(* IEC 61131-3 sources: ayran-mini-fabrika/plc/build (part 7) *)

  CASE STP OF
    0:  (* idle *)
      WANT := WORD#0;
      PUMP_REQ := FALSE;
      IF NOT WAIT_START AND (ALARMS AND ALARM_MASK) = WORD#0 THEN
        IF CIP_REQ THEN
          CIP_REQ := FALSE;
          STP := 40;
        ELSIF REQ AND NOT CIP_DUE AND NOT DI_T1_LOW THEN
          BATCH := 0;
          IF LINE_PRODUCT THEN STP := 10; ELSE STP := 20; END_IF;
        END_IF;
      END_IF;

    20: (* fill the line with product: first liquid to the drain *)
      WANT := WORD#16#0022;            (* V_PROD + V_DRAIN *)
      PUMP_REQ := TRUE;
      IF T_INWIN.Q THEN
        LINE_PRODUCT := TRUE;
        STP := 10;                     (* the route manager stops the pump and changes the route *)
      ELSIF STEP_SCANS > 2250 THEN
        ALARMS := ALARMS OR WORD#16#0200;   (* product conductivity not detected within 45 s *)
      END_IF;

    10: (* transfer to the filling tank *)
      WANT := WORD#16#0012;            (* V_PROD + V_FILL *)
      PUMP_REQ := TRUE;
      IF T_FOREIGN.Q THEN
        LINE_PRODUCT := FALSE;
        ALARMS := ALARMS OR WORD#16#0004;
      ELSIF NOT REQ OR DI_T1_LOW OR SINCE >= CIP_LIMIT OR CIP_REQ THEN
        STP := 0;
      END_IF;

    40: (* CIP preparation: empty route for the line, prove all valves closed *)
      WANT := WORD#0;
      PUMP_REQ := FALSE;
      LINE_PRODUCT := FALSE;
      CAUSTIC_IN := FALSE;
      CIP_SCANS := 0;
      MIN_T := 32000;
      MIN_F := 32000;
      FINAL_COND := 0;
      IF IW_CIP_LVL < CIP_LVL_MIN THEN
        ALARMS := ALARMS OR WORD#16#0100;
      ELSIF RSTATE = 0 AND ROUTE_OK THEN
        STP := 41;
      END_IF;

    41: (* wait for the caustic temperature *)
      WANT := WORD#0;
      PUMP_REQ := FALSE;
      IF IW_CIP_T >= CAUSTIC_SP - 50 THEN
        STP := 42;
      ELSIF STEP_TO THEN
        ALARMS := ALARMS OR WORD#16#0080;
      END_IF;

    42: (* pre-rinse: water to the drain *)
      WANT := WORD#16#0024;            (* V_WATER + V_DRAIN *)
      PUMP_REQ := TRUE;
      IF VOL >= RINSE_KG THEN
        WATER_REF := IW_COND;           (* conductivity of the inlet water: the criterion for the final rinse *)
        STP := 43;
      ELSIF STEP_TO THEN
        ALARMS := ALARMS OR WORD#16#0080;
      END_IF;

    43: (* caustic: first to the drain, to the caustic tank once caustic arrives (phase separation) *)
      PUMP_REQ := TRUE;
      IF NOT CAUSTIC_IN AND RSTATE = 0 AND IW_COND >= COND_CAUSTIC THEN CAUSTIC_IN := TRUE; END_IF;
      IF CAUSTIC_IN THEN
        WANT := WORD#16#0048;          (* V_CAUSTIC + V_CIPRET *)
      ELSE
        WANT := WORD#16#0028;          (* V_CAUSTIC + V_DRAIN *)
      END_IF;
      (* CIP record: the lowest values in the counted hold window *)
      IF HOLD_OK THEN
        IF IW_RET_T < MIN_T THEN MIN_T := IW_RET_T; END_IF;
        IF IW_FLOW < MIN_F THEN MIN_F := IW_FLOW; END_IF;
      ELSE
        MIN_T := 32000;
        MIN_F := 32000;
      END_IF;
      IF T_HOLD.Q THEN
        STP := 44;
      ELSIF STEP_TO THEN
        ALARMS := ALARMS OR WORD#16#0080;
      END_IF;

    44: (* final rinse: until no caustic is left *)
      WANT := WORD#16#0024;
      PUMP_REQ := TRUE;
      IF VOL >= RINSE_KG AND IW_COND <= WATER_REF + RINSE_MARGIN THEN
        FINAL_COND := IW_COND;
        STP := 45;
      ELSIF STEP_TO THEN
        ALARMS := ALARMS OR WORD#16#0080;
      END_IF;

    45: (* completed *)
      WANT := WORD#0;
      PUMP_REQ := FALSE;
      SINCE := 0;
      CIP_DUE := FALSE;
      ABORT_WARN := FALSE;
      CIP_RES := 1;
      CIP_DUR := CIP_SCANS / 50;
      STP := 0;
  END_CASE;
  IF STP >= 40 AND STP <= 44 AND CIP_SCANS < 30000 THEN CIP_SCANS := CIP_SCANS + 1; END_IF;
  IF CIP_RES = 2 OR CIP_RES = 3 THEN CIP_DUR := CIP_SCANS / 50; END_IF;

  (* =================== 4. Route manager =================== *)
  IF (ALARMS AND ALARM_MASK) <> WORD#0 THEN WANT := WORD#0; END_IF;
  IF WANT <> CUR AND RSTATE = 0 THEN RSTATE := 1; END_IF;
  T_ROUTE(IN := RSTATE = 1, PT := T#3s);
  T_STROKE(IN := RSTATE = 2, PT := T#1s);
  IF RSTATE = 1 THEN
    VALVES := CUR AND WANT;            (* close the ones not in the new route *)
    IF ((NOT WANT) AND WORD#16#007E AND (NOT CLOSED)) = WORD#0 THEN
      RSTATE := 2;
    ELSIF T_ROUTE.Q THEN
      ALARMS := ALARMS OR WORD#16#0008;
      RSTATE := 0;
      CUR := CUR AND WANT;
    END_IF;
  ELSIF RSTATE = 2 THEN
    VALVES := WANT;
    IF T_STROKE.Q THEN CUR := WANT; RSTATE := 0; END_IF;
  ELSE
    VALVES := CUR;
  END_IF;

  Q_P1 := PUMP_REQ AND RSTATE = 0 AND CUR = WANT AND CUR <> WORD#0 AND ROUTE_OK
          AND (ALARMS AND ALARM_MASK) = WORD#0;

  (* caustic tank thermostat (+/- 2 C), level and over-temperature interlock *)
  IF NOT ESTOP_OK OR IW_CIP_LVL < CIP_LVL_MIN OR IW_CIP_T > CAUSTIC_MAX THEN
    Q_HEAT := FALSE;
  ELSIF IW_CIP_T < CAUSTIC_SP - 20 THEN
    Q_HEAT := TRUE;
  ELSIF IW_CIP_T > CAUSTIC_SP + 20 THEN
    Q_HEAT := FALSE;
  END_IF;

  (* =================== 5. Outputs =================== *)
  WARNS := WORD#0;
  IF DI_T1_LOW THEN WARNS := WARNS OR WORD#16#0400; END_IF;
  IF CIP_DUE THEN WARNS := WARNS OR WORD#16#0800; END_IF;
  IF ABORT_WARN THEN WARNS := WARNS OR WORD#16#1000; END_IF;

  QW_DO := VALVES AND WORD#16#007E;
  IF Q_P1 THEN QW_DO := QW_DO OR WORD#16#0001; END_IF;
  IF Q_HEAT THEN QW_DO := QW_DO OR WORD#16#0080; END_IF;
  IF STP >= 40 THEN QW_DO := QW_DO OR WORD#16#0100; END_IF;

  IF (ALARMS AND WORD#16#0001) <> WORD#0 THEN
    QW_STATE := 11;
  ELSIF (ALARMS AND ALARM_MASK) <> WORD#0 THEN
    QW_STATE := 10;
  ELSIF STP = 0 AND CIP_DUE THEN
    QW_STATE := 9;
  ELSIF STP = 0 THEN
    QW_STATE := 0;
  ELSIF (STP = 10 OR STP = 20) AND RSTATE <> 0 THEN
    QW_STATE := 3;
  ELSIF STP = 10 THEN
    QW_STATE := 1;
  ELSIF STP = 20 THEN
    QW_STATE := 2;
  ELSE
    QW_STATE := STP - 36;             (* 40..44 -> 4..8 *)
  END_IF;

  QW_ALARM    := ALARMS OR WARNS;
  QW_STEP_T   := STEP_SCANS / 50;
  QW_SINCE    := SINCE;
  QW_BATCH    := BATCH;
  QW_CIP_RES  := CIP_RES;
  IF MIN_T = 32000 THEN QW_CIP_MINT := 0; ELSE QW_CIP_MINT := MIN_T; END_IF;
  IF MIN_F = 32000 THEN QW_CIP_MINF := 0; ELSE QW_CIP_MINF := MIN_F; END_IF;
  QW_CIP_COND := FINAL_COND;
  QW_CIP_DUR  := CIP_DUR;
  TRANSFERRING := STP = 10 AND Q_P1;
  QW_STATUS := WORD#0;
  IF WAIT_START THEN QW_STATUS := WORD#16#0080; END_IF;
  IF WAIT_START OR NOT IO_READY THEN
    QW_DO := WORD#0;
    Q_HEAT := FALSE; Q_P1 := FALSE;
  END_IF;
END_FUNCTION_BLOCK

PROGRAM Proses
  VAR
    (* --- blok 0: Fabrika --- *)
    FAB_IW_DI        AT %IW100 : WORD;  (* Fabrika paneli girisleri (bit paketli) *)
    FAB_IW_MAPVER    AT %IW101 : INT;  (* Sinyal haritasi surumu *)
    FAB_IW_SIM_HB    AT %IW102 : INT;  (* Simulator kalp atisi (100 ms) *)
    FAB_QW_DO        AT %QW100 : WORD;  (* Fabrika cikislari (bit paketli) *)
    FAB_QW_PLC_HB    AT %QW101 : INT;  (* Proses PLC (ya da tek PLC) kalp atisi (her tarama) *)
    FAB_QW_STATE     AT %QW102 : INT;  (* Fabrika durumu *)
    FAB_QW_ALARM     AT %QW103 : WORD;  (* Fabrika alarm ozeti *)
    (* --- blok 1: Dolum-kapama --- *)
    DOL_IW_DI        AT %IW116 : WORD;  (* Dijital girisler (bit paketli) *)
    DOL_IW_FILL      AT %IW117 : INT;  (* Dolum terazisi (net) *)
    DOL_IW_TANK      AT %IW118 : INT;  (* Dolum tanki seviyesi *)
    DOL_IW_TEMP      AT %IW119 : INT;  (* Kapama kafasi sicakligi *)
    DOL_IW_CHECK     AT %IW120 : INT;  (* Kontrol tartisi (brut) *)
    DOL_QW_DO        AT %QW116 : WORD;  (* Dijital cikislar (bit paketli) *)
    DOL_QW_STATE     AT %QW117 : INT;  (* Makine modu *)
    DOL_QW_ALARM     AT %QW118 : WORD;  (* Alarm kelimesi *)
    DOL_QW_GOOD      AT %QW119 : INT;  (* Saglam bardak sayaci *)
    DOL_QW_REJECT    AT %QW120 : INT;  (* Red sayaci *)
    DOL_QW_STATUS    AT %QW121 : WORD;  (* Durum bitleri (bit 7: yeniden basladi, START bekliyor) *)
    (* --- blok 2: Tank ve transfer --- *)
    TNK_IW_DI        AT %IW132 : WORD;  (* Dijital girisler (bit paketli) *)
    TNK_IW_T1_LVL    AT %IW133 : INT;  (* Uretim tanki T1 seviyesi *)
    TNK_IW_FLOW      AT %IW134 : INT;  (* Debimetre FT1 *)
    TNK_IW_TOTAL     AT %IW135 : INT;  (* Debimetre toplayici (30000'de sifirlanir) *)
    TNK_IW_COND      AT %IW136 : INT;  (* Hat iletkenligi QT1 (25 ?C'ye duzeltilmis) *)
    TNK_IW_RET_T     AT %IW137 : INT;  (* Hat donus sicakligi TT1 *)
    TNK_IW_CIP_T     AT %IW138 : INT;  (* Kostik tanki sicakligi TT2 *)
    TNK_IW_CIP_LVL   AT %IW139 : INT;  (* Kostik tanki seviyesi *)
    TNK_QW_DO        AT %QW132 : WORD;  (* Dijital cikislar (bit paketli) *)
    TNK_QW_STATE     AT %QW133 : INT;  (* Istasyon durumu *)
    TNK_QW_ALARM     AT %QW134 : WORD;  (* Alarm kelimesi *)
    TNK_QW_STEP_T    AT %QW135 : INT;  (* Adim suresi *)
    TNK_QW_SINCE     AT %QW136 : INT;  (* Son CIP'ten beri aktarilan *)
    TNK_QW_BATCH     AT %QW137 : INT;  (* Bu aktarimda aktarilan *)
    TNK_QW_CIP_RES   AT %QW138 : INT;  (* Son CIP sonucu (0 yok, 1 basarili, 2 iptal, 3 basarisiz) *)
    TNK_QW_CIP_MINT  AT %QW139 : INT;  (* Son CIP: tutma sirasinda en dusuk donus sicakligi *)
    TNK_QW_CIP_MINF  AT %QW140 : INT;  (* Son CIP: tutma sirasinda en dusuk debi *)
    TNK_QW_CIP_COND  AT %QW141 : INT;  (* Son CIP: son durulama iletkenligi *)
    TNK_QW_CIP_DUR   AT %QW142 : INT;  (* Son CIP: toplam sure *)
    TNK_QW_STATUS    AT %QW143 : WORD;  (* Durum bitleri (bit 7: yeniden basladi, START bekliyor) *)
    TNK_COMMISSION AT %MW0 : WORD;
  END_VAR

  VAR
    PB_START    : BOOL;   (* factory panel *)
    PB_STOP_OK  : BOOL;
    PB_ESTOP_OK : BOOL;
    PB_RESET    : BOOL;
    FIRST_SCAN  : BOOL := TRUE;
    RESTART     : BOOL;
    IO_READY    : BOOL;   (* first data arrived from the simulator with the correct version *)
    COMM_FAULT  : BOOL;
    SIM_HB_LAST : INT;
    PLC_HB      : INT;
    T_SIMHB     : TON;
    DOLUM       : FB_Dolum;
    TANK        : FB_Tank;
  END_VAR

  (* =================== 1. Factory panel =================== *)
  PB_START    := (FAB_IW_DI AND WORD#16#0001) <> WORD#0;
  PB_STOP_OK  := (FAB_IW_DI AND WORD#16#0002) <> WORD#0;
  PB_ESTOP_OK := (FAB_IW_DI AND WORD#16#0004) <> WORD#0;
  PB_RESET    := (FAB_IW_DI AND WORD#16#0008) <> WORD#0;

  (* =================== 2. Communication watchdog =================== *)
  (* communication fault if the simulator heartbeat does not change for 2 s *)
  T_SIMHB(IN := (FAB_IW_SIM_HB = SIM_HB_LAST), PT := T#2s);
  SIM_HB_LAST := FAB_IW_SIM_HB;
  COMM_FAULT := T_SIMHB.Q;
  (* inputs are invalid until the first data arrives and the map version matches *)
  IF FAB_IW_SIM_HB <> 0 AND FAB_IW_MAPVER = 7 THEN IO_READY := TRUE; END_IF;

  RESTART := FIRST_SCAN AND IO_READY;
  IF RESTART THEN FIRST_SCAN := FALSE; END_IF;

  (* PLC heartbeat: the simulator watches it and switches off this PLC's outputs if the program stops *)
  PLC_HB := PLC_HB + 1;
  IF PLC_HB > 30000 THEN PLC_HB := 0; END_IF;

  (* =================== Fill-and-seal =================== *)
  DOLUM(START := PB_START, STOP_OK := PB_STOP_OK, ESTOP_OK := PB_ESTOP_OK, RESET := PB_RESET,
        RESTART := RESTART, IO_READY := IO_READY, COMM_FAULT := COMM_FAULT,
        IW_DI := DOL_IW_DI, IW_FILL := DOL_IW_FILL, IW_TANK := DOL_IW_TANK,
        IW_TEMP := DOL_IW_TEMP, IW_CHECK := DOL_IW_CHECK);
  DOL_QW_DO     := DOLUM.QW_DO;
  DOL_QW_STATE  := DOLUM.QW_STATE;
  DOL_QW_ALARM  := DOLUM.QW_ALARM;
  DOL_QW_GOOD   := DOLUM.QW_GOOD;
  DOL_QW_REJECT := DOLUM.QW_REJECT;
  DOL_QW_STATUS := DOLUM.QW_STATUS;

  (* handshake: the filling machine requests product, the tank station transfers it (same PLC) *)
  TANK(START := PB_START, TNK_COMMISSION := TNK_COMMISSION, ESTOP_OK := PB_ESTOP_OK, RESET := PB_RESET, RESTART := RESTART, IO_READY := IO_READY, COMM_FAULT := COMM_FAULT,
       REQ := DOLUM.PRODUCT_REQ,
       IW_DI := TNK_IW_DI, IW_T1_LVL := TNK_IW_T1_LVL, IW_FLOW := TNK_IW_FLOW, IW_TOTAL := TNK_IW_TOTAL,
       IW_COND := TNK_IW_COND, IW_RET_T := TNK_IW_RET_T, IW_CIP_T := TNK_IW_CIP_T, IW_CIP_LVL := TNK_IW_CIP_LVL);
  TNK_QW_DO       := TANK.QW_DO;
  TNK_QW_STATE    := TANK.QW_STATE;
  TNK_QW_ALARM    := TANK.QW_ALARM;
  TNK_QW_STEP_T   := TANK.QW_STEP_T;
  TNK_QW_SINCE    := TANK.QW_SINCE;
  TNK_QW_BATCH    := TANK.QW_BATCH;
  TNK_QW_CIP_RES  := TANK.QW_CIP_RES;
  TNK_QW_CIP_MINT := TANK.QW_CIP_MINT;
  TNK_QW_CIP_MINF := TANK.QW_CIP_MINF;
  TNK_QW_CIP_COND := TANK.QW_CIP_COND;
  TNK_QW_CIP_DUR  := TANK.QW_CIP_DUR;
  TNK_QW_STATUS := TANK.QW_STATUS;

  (* =================== Factory summary (block 0) =================== *)
  FAB_QW_PLC_HB := PLC_HB;
  IF DOLUM.RUNNING THEN FAB_QW_DO := WORD#16#0001; ELSE FAB_QW_DO := WORD#0; END_IF;
  FAB_QW_STATE := DOLUM.QW_STATE;
  FAB_QW_ALARM := DOLUM.QW_ALARM OR TANK.QW_ALARM;
END_PROGRAM

CONFIGURATION Config0
  RESOURCE Res0 ON PLC
    TASK task0(INTERVAL := T#20ms, PRIORITY := 0);
    PROGRAM instance0 WITH task0 : Proses;
  END_RESOURCE
END_CONFIGURATION
